(* IEC 61131-3 sources: plc_generation_empirical_study/datasets/_archive/pre_native_plcverif_20260810/tasks/C10_E01_master_follower_coordination, 2 files *)

(* ---- interface.st ---- *)
FUNCTION_BLOCK C10_E01_master_follower_coordination
VAR_INPUT
    RunRequest : BOOL;
    MasterReady : BOOL;
    FollowerReady : BOOL;
END_VAR
VAR_OUTPUT
    MasterRun : BOOL;
    FollowerRun : BOOL;
END_VAR
END_FUNCTION_BLOCK

(* ---- reference.st ---- *)
FUNCTION_BLOCK C10_E01_master_follower_coordination
VAR_INPUT
    RunRequest : BOOL;
    MasterReady : BOOL;
    FollowerReady : BOOL;
END_VAR
VAR_OUTPUT
    MasterRun : BOOL;
    FollowerRun : BOOL;
END_VAR

MasterRun := RunRequest AND MasterReady;
FollowerRun := RunRequest AND MasterRun AND FollowerReady;

END_FUNCTION_BLOCK
